// TIA Portal V19 export
FUNCTION "G120XA_DATA_MAPPING" : Void   // FC5, LAD
{ S7_Optimized_Access := 'TRUE' }
// stored: SetENOAutomatically false
BEGIN

REGION Network 1: COLD_SKID_CP01
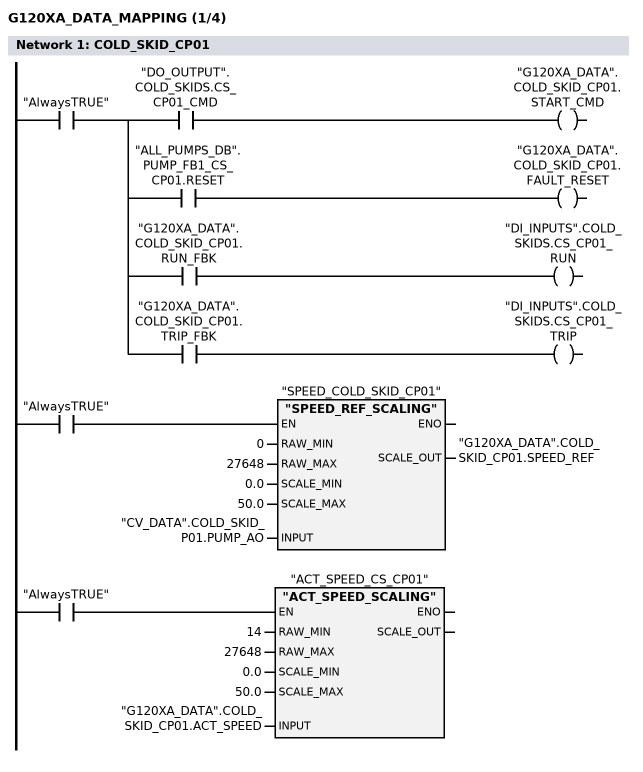
   RUNG wire#powerrail
      Contact( "AlwaysTRUE" )
      wire#w1
      Contact( "DO_OUTPUT".COLD_SKIDS.CS_CP01_CMD )
      Coil( "G120XA_DATA".COLD_SKID_CP01.START_CMD )
   END_RUNG
   RUNG wire#w1
      Contact( "ALL_PUMPS_DB".PUMP_FB1_CS_CP01.RESET )
      Coil( "G120XA_DATA".COLD_SKID_CP01.FAULT_RESET )
   END_RUNG
   RUNG wire#w1
      Contact( "G120XA_DATA".COLD_SKID_CP01.RUN_FBK )
      Coil( "DI_INPUTS".COLD_SKIDS.CS_CP01_RUN )
   END_RUNG
   RUNG wire#w1
      Contact( "G120XA_DATA".COLD_SKID_CP01.TRIP_FBK )
      Coil( "DI_INPUTS".COLD_SKIDS.CS_CP01_TRIP )
   END_RUNG
   RUNG wire#powerrail
      Contact( "AlwaysTRUE" )
      "SPEED_COLD_SKID_CP01"(RAW_MIN := 0, RAW_MAX := 27648, SCALE_MIN := 0.0, SCALE_MAX := 50.0, INPUT := "CV_DATA".COLD_SKID_P01.PUMP_AO, SCALE_OUT => "G120XA_DATA".COLD_SKID_CP01.SPEED_REF)
   END_RUNG
   RUNG wire#powerrail
      Contact( "AlwaysTRUE" )
      "ACT_SPEED_CS_CP01"(RAW_MIN := 14, RAW_MAX := 27648, SCALE_MIN := 0.0, SCALE_MAX := 50.0, INPUT := "G120XA_DATA".COLD_SKID_CP01.ACT_SPEED, SCALE_OUT =>)
   END_RUNG
   // the same network as SCL:
   "G120XA_DATA".COLD_SKID_CP01.START_CMD := "AlwaysTRUE" AND "DO_OUTPUT".COLD_SKIDS.CS_CP01_CMD;
   "G120XA_DATA".COLD_SKID_CP01.FAULT_RESET := "AlwaysTRUE" AND "ALL_PUMPS_DB".PUMP_FB1_CS_CP01.RESET;
   "DI_INPUTS".COLD_SKIDS.CS_CP01_RUN := "AlwaysTRUE" AND "G120XA_DATA".COLD_SKID_CP01.RUN_FBK;
   "DI_INPUTS".COLD_SKIDS.CS_CP01_TRIP := "AlwaysTRUE" AND "G120XA_DATA".COLD_SKID_CP01.TRIP_FBK;
   IF "AlwaysTRUE" THEN
       "SPEED_COLD_SKID_CP01"(RAW_MIN := 0,   // "SPEED_REF_SCALING"
                              RAW_MAX := 27648,
                              SCALE_MIN := 0.0,
                              SCALE_MAX := 50.0,
                              INPUT := "CV_DATA".COLD_SKID_P01.PUMP_AO,
                              SCALE_OUT => "G120XA_DATA".COLD_SKID_CP01.SPEED_REF);
   END_IF;
   IF "AlwaysTRUE" THEN
       "ACT_SPEED_CS_CP01"(RAW_MIN := 14,   // "ACT_SPEED_SCALING"
                           RAW_MAX := 27648,
                           SCALE_MIN := 0.0,
                           SCALE_MAX := 50.0,
                           INPUT := "G120XA_DATA".COLD_SKID_CP01.ACT_SPEED);
   END_IF;
END_REGION

REGION Network 2: COLD_SKID_CP02
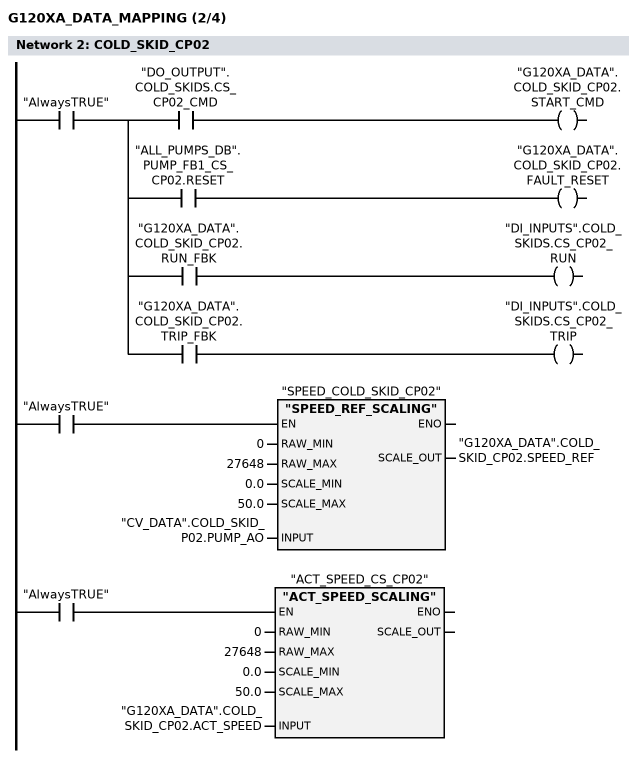
   RUNG wire#powerrail
      Contact( "AlwaysTRUE" )
      wire#w1
      Contact( "DO_OUTPUT".COLD_SKIDS.CS_CP02_CMD )
      Coil( "G120XA_DATA".COLD_SKID_CP02.START_CMD )
   END_RUNG
   RUNG wire#w1
      Contact( "ALL_PUMPS_DB".PUMP_FB1_CS_CP02.RESET )
      Coil( "G120XA_DATA".COLD_SKID_CP02.FAULT_RESET )
   END_RUNG
   RUNG wire#w1
      Contact( "G120XA_DATA".COLD_SKID_CP02.RUN_FBK )
      Coil( "DI_INPUTS".COLD_SKIDS.CS_CP02_RUN )
   END_RUNG
   RUNG wire#w1
      Contact( "G120XA_DATA".COLD_SKID_CP02.TRIP_FBK )
      Coil( "DI_INPUTS".COLD_SKIDS.CS_CP02_TRIP )
   END_RUNG
   RUNG wire#powerrail
      Contact( "AlwaysTRUE" )
      "SPEED_COLD_SKID_CP02"(RAW_MIN := 0, RAW_MAX := 27648, SCALE_MIN := 0.0, SCALE_MAX := 50.0, INPUT := "CV_DATA".COLD_SKID_P02.PUMP_AO, SCALE_OUT => "G120XA_DATA".COLD_SKID_CP02.SPEED_REF)
   END_RUNG
   RUNG wire#powerrail
      Contact( "AlwaysTRUE" )
      "ACT_SPEED_CS_CP02"(RAW_MIN := 0, RAW_MAX := 27648, SCALE_MIN := 0.0, SCALE_MAX := 50.0, INPUT := "G120XA_DATA".COLD_SKID_CP02.ACT_SPEED, SCALE_OUT =>)
   END_RUNG
   // the same network as SCL:
   "G120XA_DATA".COLD_SKID_CP02.START_CMD := "AlwaysTRUE" AND "DO_OUTPUT".COLD_SKIDS.CS_CP02_CMD;
   "G120XA_DATA".COLD_SKID_CP02.FAULT_RESET := "AlwaysTRUE" AND "ALL_PUMPS_DB".PUMP_FB1_CS_CP02.RESET;
   "DI_INPUTS".COLD_SKIDS.CS_CP02_RUN := "AlwaysTRUE" AND "G120XA_DATA".COLD_SKID_CP02.RUN_FBK;
   "DI_INPUTS".COLD_SKIDS.CS_CP02_TRIP := "AlwaysTRUE" AND "G120XA_DATA".COLD_SKID_CP02.TRIP_FBK;
   IF "AlwaysTRUE" THEN
       "SPEED_COLD_SKID_CP02"(RAW_MIN := 0,   // "SPEED_REF_SCALING"
                              RAW_MAX := 27648,
                              SCALE_MIN := 0.0,
                              SCALE_MAX := 50.0,
                              INPUT := "CV_DATA".COLD_SKID_P02.PUMP_AO,
                              SCALE_OUT => "G120XA_DATA".COLD_SKID_CP02.SPEED_REF);
   END_IF;
   IF "AlwaysTRUE" THEN
       "ACT_SPEED_CS_CP02"(RAW_MIN := 0,   // "ACT_SPEED_SCALING"
                           RAW_MAX := 27648,
                           SCALE_MIN := 0.0,
                           SCALE_MAX := 50.0,
                           INPUT := "G120XA_DATA".COLD_SKID_CP02.ACT_SPEED);
   END_IF;
END_REGION

REGION Network 3: COLD_SKID_CP01
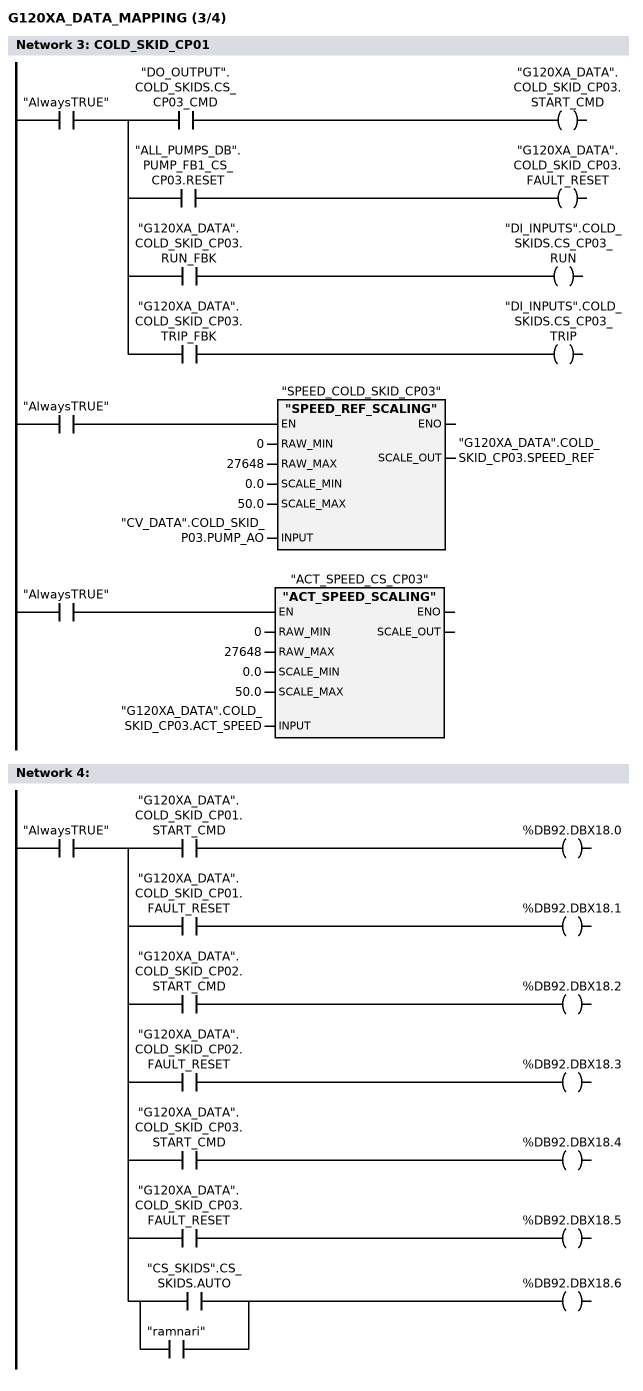
   RUNG wire#powerrail
      Contact( "AlwaysTRUE" )
      wire#w1
      Contact( "DO_OUTPUT".COLD_SKIDS.CS_CP03_CMD )
      Coil( "G120XA_DATA".COLD_SKID_CP03.START_CMD )
   END_RUNG
   RUNG wire#w1
      Contact( "ALL_PUMPS_DB".PUMP_FB1_CS_CP03.RESET )
      Coil( "G120XA_DATA".COLD_SKID_CP03.FAULT_RESET )
   END_RUNG
   RUNG wire#w1
      Contact( "G120XA_DATA".COLD_SKID_CP03.RUN_FBK )
      Coil( "DI_INPUTS".COLD_SKIDS.CS_CP03_RUN )
   END_RUNG
   RUNG wire#w1
      Contact( "G120XA_DATA".COLD_SKID_CP03.TRIP_FBK )
      Coil( "DI_INPUTS".COLD_SKIDS.CS_CP03_TRIP )
   END_RUNG
   RUNG wire#powerrail
      Contact( "AlwaysTRUE" )
      "SPEED_COLD_SKID_CP03"(RAW_MIN := 0, RAW_MAX := 27648, SCALE_MIN := 0.0, SCALE_MAX := 50.0, INPUT := "CV_DATA".COLD_SKID_P03.PUMP_AO, SCALE_OUT => "G120XA_DATA".COLD_SKID_CP03.SPEED_REF)
   END_RUNG
   RUNG wire#powerrail
      Contact( "AlwaysTRUE" )
      "ACT_SPEED_CS_CP03"(RAW_MIN := 0, RAW_MAX := 27648, SCALE_MIN := 0.0, SCALE_MAX := 50.0, INPUT := "G120XA_DATA".COLD_SKID_CP03.ACT_SPEED, SCALE_OUT =>)
   END_RUNG
   // the same network as SCL:
   "G120XA_DATA".COLD_SKID_CP03.START_CMD := "AlwaysTRUE" AND "DO_OUTPUT".COLD_SKIDS.CS_CP03_CMD;
   "G120XA_DATA".COLD_SKID_CP03.FAULT_RESET := "AlwaysTRUE" AND "ALL_PUMPS_DB".PUMP_FB1_CS_CP03.RESET;
   "DI_INPUTS".COLD_SKIDS.CS_CP03_RUN := "AlwaysTRUE" AND "G120XA_DATA".COLD_SKID_CP03.RUN_FBK;
   "DI_INPUTS".COLD_SKIDS.CS_CP03_TRIP := "AlwaysTRUE" AND "G120XA_DATA".COLD_SKID_CP03.TRIP_FBK;
   IF "AlwaysTRUE" THEN
       "SPEED_COLD_SKID_CP03"(RAW_MIN := 0,   // "SPEED_REF_SCALING"
                              RAW_MAX := 27648,
                              SCALE_MIN := 0.0,
                              SCALE_MAX := 50.0,
                              INPUT := "CV_DATA".COLD_SKID_P03.PUMP_AO,
                              SCALE_OUT => "G120XA_DATA".COLD_SKID_CP03.SPEED_REF);
   END_IF;
   IF "AlwaysTRUE" THEN
       "ACT_SPEED_CS_CP03"(RAW_MIN := 0,   // "ACT_SPEED_SCALING"
                           RAW_MAX := 27648,
                           SCALE_MIN := 0.0,
                           SCALE_MAX := 50.0,
                           INPUT := "G120XA_DATA".COLD_SKID_CP03.ACT_SPEED);
   END_IF;
END_REGION

REGION Network 4
   RUNG wire#powerrail
      Contact( "AlwaysTRUE" )
      wire#w1
      Contact( "G120XA_DATA".COLD_SKID_CP01.START_CMD )
      Coil( %DB92.DBX18.0 )
   END_RUNG
   RUNG wire#w1
      Contact( "G120XA_DATA".COLD_SKID_CP01.FAULT_RESET )
      Coil( %DB92.DBX18.1 )
   END_RUNG
   RUNG wire#w1
      Contact( "G120XA_DATA".COLD_SKID_CP02.START_CMD )
      Coil( %DB92.DBX18.2 )
   END_RUNG
   RUNG wire#w1
      Contact( "G120XA_DATA".COLD_SKID_CP02.FAULT_RESET )
      Coil( %DB92.DBX18.3 )
   END_RUNG
   RUNG wire#w1
      Contact( "G120XA_DATA".COLD_SKID_CP03.START_CMD )
      Coil( %DB92.DBX18.4 )
   END_RUNG
   RUNG wire#w1
      Contact( "G120XA_DATA".COLD_SKID_CP03.FAULT_RESET )
      Coil( %DB92.DBX18.5 )
   END_RUNG
   RUNG wire#w1
      Contact( "CS_SKIDS".CS_SKIDS.AUTO )
      wire#w2
      Coil( %DB92.DBX18.6 )
   END_RUNG
   RUNG wire#w1
      Contact( "ramnari" )
   END_RUNG wire#w2
   // the same network as SCL:
   %DB92.DBX18.0 := "AlwaysTRUE" AND "G120XA_DATA".COLD_SKID_CP01.START_CMD;
   %DB92.DBX18.1 := "AlwaysTRUE" AND "G120XA_DATA".COLD_SKID_CP01.FAULT_RESET;
   %DB92.DBX18.2 := "AlwaysTRUE" AND "G120XA_DATA".COLD_SKID_CP02.START_CMD;
   %DB92.DBX18.3 := "AlwaysTRUE" AND "G120XA_DATA".COLD_SKID_CP02.FAULT_RESET;
   %DB92.DBX18.4 := "AlwaysTRUE" AND "G120XA_DATA".COLD_SKID_CP03.START_CMD;
   %DB92.DBX18.5 := "AlwaysTRUE" AND "G120XA_DATA".COLD_SKID_CP03.FAULT_RESET;
   %DB92.DBX18.6 := "AlwaysTRUE" AND ("CS_SKIDS".CS_SKIDS.AUTO OR "ramnari");
END_REGION

REGION Network 5
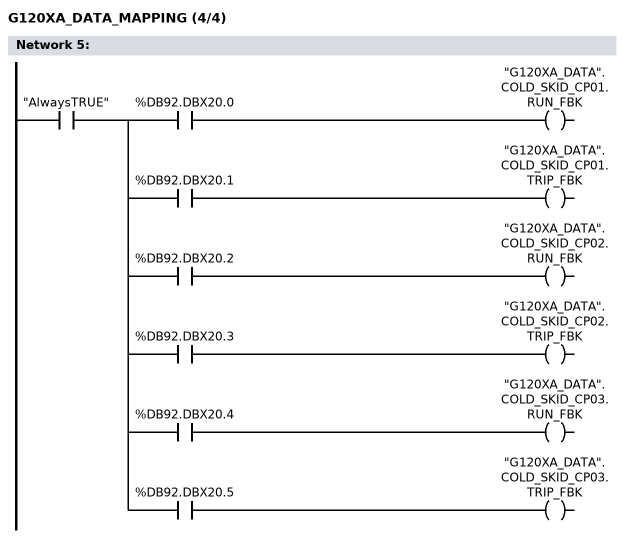
   RUNG wire#powerrail
      Contact( "AlwaysTRUE" )
      wire#w1
      Contact( %DB92.DBX20.0 )
      Coil( "G120XA_DATA".COLD_SKID_CP01.RUN_FBK )
   END_RUNG
   RUNG wire#w1
      Contact( %DB92.DBX20.1 )
      Coil( "G120XA_DATA".COLD_SKID_CP01.TRIP_FBK )
   END_RUNG
   RUNG wire#w1
      Contact( %DB92.DBX20.2 )
      Coil( "G120XA_DATA".COLD_SKID_CP02.RUN_FBK )
   END_RUNG
   RUNG wire#w1
      Contact( %DB92.DBX20.3 )
      Coil( "G120XA_DATA".COLD_SKID_CP02.TRIP_FBK )
   END_RUNG
   RUNG wire#w1
      Contact( %DB92.DBX20.4 )
      Coil( "G120XA_DATA".COLD_SKID_CP03.RUN_FBK )
   END_RUNG
   RUNG wire#w1
      Contact( %DB92.DBX20.5 )
      Coil( "G120XA_DATA".COLD_SKID_CP03.TRIP_FBK )
   END_RUNG
   // the same network as SCL:
   "G120XA_DATA".COLD_SKID_CP01.RUN_FBK := "AlwaysTRUE" AND %DB92.DBX20.0;
   "G120XA_DATA".COLD_SKID_CP01.TRIP_FBK := "AlwaysTRUE" AND %DB92.DBX20.1;
   "G120XA_DATA".COLD_SKID_CP02.RUN_FBK := "AlwaysTRUE" AND %DB92.DBX20.2;
   "G120XA_DATA".COLD_SKID_CP02.TRIP_FBK := "AlwaysTRUE" AND %DB92.DBX20.3;
   "G120XA_DATA".COLD_SKID_CP03.RUN_FBK := "AlwaysTRUE" AND %DB92.DBX20.4;
   "G120XA_DATA".COLD_SKID_CP03.TRIP_FBK := "AlwaysTRUE" AND %DB92.DBX20.5;
END_REGION
END_FUNCTION
